Yaskawa INFORM job: LONGPRO5.JBI

/JOB
//NAME LONGPRO5
//POS
///NPOS 3,0,0,0,0,0
///TOOL 9
///POSTYPE PULSE
///PULSE
C00000=20480,-10240,0,-34475,0,-8704,22983
C00001=0,-10240,0,-34475,0,0,22983
C00002=20480,-10240,0,-34475,0,-8704,22983
//INST
<volatile>
///COMM Generated using RoboDK
///ATTR SC,RW
///GROUP1 RB1
NOP
MOVJ C00000 VJ=50.00
MOVJ C00001 VJ=50.00
MOVJ C00002 VJ=50.00
END
